ABB RAPID module: TgtProg.mod

MODULE MainModule

GLOBAL Proc main()
    wobj16.x = 1.23456
    wobj16.y = 2.000
    wobj16.z = 3.000
    wobj16.q1 = 0.997151
    wobj16.q2 = 0.050734
    wobj16.q3 = 0.045358
    wobj16.q4 = 0.032537
    wobj16.x = -0.0
    wobj16.y = 2.000
    wobj16.z = 3.000
    wobj16.q1 = 0.997151
    wobj16.q2 = 0.050734
    wobj16.q3 = 0.045358
    wobj16.q4 = 0.032537
    wobj16.x = 12345678.9
    wobj16.y = 2.000
    wobj16.z = 3.000
    wobj16.q1 = 0.997151
    wobj16.q2 = 0.050734
    wobj16.q3 = 0.045358
    wobj16.q4 = 0.032537
    tool03.x = 1.235
    tool03.y = 2.000
    tool03.z = 3.000
    tool03.q1 = 0.997151
    tool03.q2 = 0.050734
    tool03.q3 = 0.045358
    tool03.q4 = 0.032537
EndProc
EndModule
